FUNCTION_BLOCK FB_ConveyorProperties
VAR
    requested : BOOL;
    runningState : BOOL;
    resetStartup : BOOL;
    configuredDelay : TIME := T#1s;
    speed : LREAL := 0.5;
    count : UDINT;
    alarmText : STRING(80);
END_VAR

(* The program invokes methods explicitly. *)

METHOD PUBLIC Start
VAR_INPUT
    delay : TIME := T#1s;
END_VAR
THIS^.configuredDelay := delay;
THIS^.requested := TRUE;
END_METHOD

METHOD PUBLIC Stop
THIS^.requested := FALSE;
THIS^.runningState := FALSE;
THIS^.resetStartup := TRUE;
THIS^.alarmText := 'Stopped';
END_METHOD

METHOD PUBLIC Reset
THIS^.count := 0;
END_METHOD

METHOD PUBLIC Update : UDINT
VAR_INPUT
    guardClosed : BOOL;
    stopRequested : BOOL := FALSE;
    sensor : BOOL := FALSE;
END_VAR
VAR_INST
    startup : TON;
    productEdge : R_TRIG;
    updates : UDINT;
END_VAR
(* All three VAR_INST variables belong to this conveyor and this method. *)
updates := updates + 1;
IF stopRequested OR NOT guardClosed THEN
    THIS^.Stop();
END_IF;
IF THIS^.resetStartup THEN
    startup(IN := FALSE, PT := THIS^.configuredDelay);
    THIS^.resetStartup := FALSE;
END_IF;
startup(IN := THIS^.requested, PT := THIS^.configuredDelay);
THIS^.runningState := startup.Q;
(* Sample while stopped too, so restart cannot manufacture an edge. *)
productEdge(CLK := sensor);
IF THIS^.runningState AND productEdge.Q THEN
    THIS^.count := THIS^.count + 1;
END_IF;
IF NOT guardClosed THEN
    THIS^.alarmText := 'Guard open';
ELSIF stopRequested THEN
    THIS^.alarmText := 'Stopped';
ELSIF THIS^.requested AND NOT THIS^.runningState THEN
    THIS^.alarmText := 'Starting';
ELSE
    THIS^.alarmText := '';
END_IF;
Update := updates;
END_METHOD

PROPERTY PUBLIC SpeedSetpoint : LREAL
GET
SpeedSetpoint := THIS^.speed;
END_GET
SET
(* The assigned property value is available in the local SpeedSetpoint slot. *)
IF SpeedSetpoint < 0.0 THEN
    THIS^.speed := 0.0;
ELSIF SpeedSetpoint > 1.0 THEN
    THIS^.speed := 1.0;
ELSE
    THIS^.speed := SpeedSetpoint;
END_IF;
END_SET
END_PROPERTY

PROPERTY PUBLIC Running : BOOL
GET
Running := THIS^.runningState;
END_GET
END_PROPERTY

PROPERTY PUBLIC ActiveSpeed : LREAL
GET
IF THIS^.Running THEN
    ActiveSpeed := THIS^.SpeedSetpoint;
ELSE
    ActiveSpeed := 0.0;
END_IF;
END_GET
END_PROPERTY

PROPERTY PUBLIC ProductCount : UDINT
GET
ProductCount := THIS^.count;
END_GET
END_PROPERTY

PROPERTY PUBLIC Alarm : STRING(80)
GET
Alarm := THIS^.alarmText;
END_GET
END_PROPERTY

END_FUNCTION_BLOCK

(* stored: Version 1.1.0.1, ProductVersion 3.1 *)
